SUBAPPLICATION mapping_DataPanel (* Subapplication Type *)
  (* Standard: 61499-2 *)
  (* Version 1.0, 2023-01-29, Franz *)
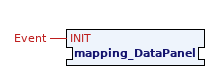
  EVENT_INPUT
    INIT;
  END_EVENT
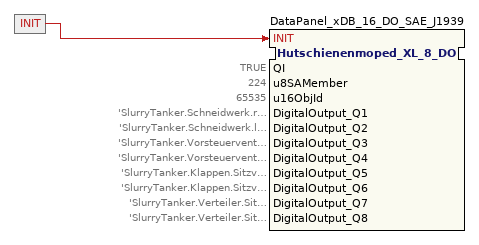
  FBS
    DataPanel_xDB_16_DO_SAE_J1939 : Hutschienenmoped_XL_8_DO(QI := TRUE, u8SAMember := 224, u16ObjId := 65535, DigitalOutput_Q1 := 'SlurryTanker.Schneidwerk.rechtslauf', DigitalOutput_Q2 := 'SlurryTanker.Schneidwerk.linkslauf', DigitalOutput_Q3 := 'SlurryTanker.Vorsteuerventil_2A.QX', DigitalOutput_Q4 := 'SlurryTanker.Vorsteuerventil_2B.QX', DigitalOutput_Q5 := 'SlurryTanker.Klappen.Sitzventile.QXA', DigitalOutput_Q6 := 'SlurryTanker.Klappen.Sitzventile.QXB', DigitalOutput_Q7 := 'SlurryTanker.Verteiler.Sitzventile.QXA', DigitalOutput_Q8 := 'SlurryTanker.Verteiler.Sitzventile.QXB');
  END_FBS
  EVENT_CONNECTIONS
    INIT TO DataPanel_xDB_16_DO_SAE_J1939.INIT;
  END_CONNECTIONS
END_SUBAPPLICATION
